Fanuc KAREL source: kb00023.KL

-- PROVISIONAL review KL for V1013-1; original PC SHA256 f590d3276f3f32f3e88922adc0d481ff6561b01a1212fb5bc6264c8695096b18
-- Incomplete behavior may be omitted. Consult companion uncertainty JSON. Do not deploy.
PROGRAM KB00023
%NOLOCKGROUP
BEGIN
  -- UNRESOLVED_PC offsets 5-12; opcodes 9D,23
  -- UNRESOLVED_PC offsets 17-24; opcodes 9D,23
  -- UNRESOLVED_PC offsets 29-45; opcodes 27,22,22,31
  -- UNRESOLVED_PC offsets 50-54; opcodes 7F
END KB00023
